FUNCTION_BLOCK SKILL_Merge (* Where the two branches of a decision meet again: either branch's end goes on. Technical: Where the branches of a decision meet: EI1 or EI2 gives EO *)
  (* Standard: 61499-2 *)
  (* Version 0.1, 2026-09-28, Project contributors, AAU Smart Production Lab *)
  PACKAGE modlib;
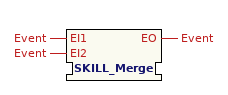
  EVENT_INPUT
    EI1; (* The first branch of the decision is done *)
    EI2; (* The second branch is done, or there was none to run *)
  END_EVENT
  EVENT_OUTPUT
    EO; (* The decision is done: the next step goes on *)
  END_EVENT
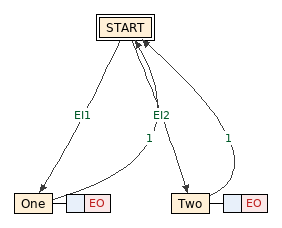
  EC_STATES
    START;
    One : -> EO;
    Two : -> EO;
  END_STATES
  EC_TRANSITIONS
    START TO One := EI1;
    START TO Two := EI2;
    One TO START := 1;
    Two TO START := 1;
  END_TRANSITIONS
END_FUNCTION_BLOCK
